// TIA Portal V20 export
// export: Created 2026-10-12T15:48:35.0909134Z, ExportSetting WithDefaults, DisplayName Totally Integrated Automation Portal, DisplayVersion V20, DisplayName TIA Portal Openness, DisplayVersion V20, DisplayName TIA Portal Teamcenter Gateway, DisplayVersion V20, DisplayName TIA Portal Version Control Interface, DisplayVersion V20, DisplayName SINAMICS Startdrive Advanced, DisplayVersion V20 SP1 Update 2, DisplayName SINAMICS Startdrive G110M, G120, G120C, G120D, G120P, G115D, DisplayVersion V20 SP1 Update 2, DisplayName SINAMICS Startdrive G130, G150, S120, S150, SINAMICS MV, G220, S200, S210, DisplayVersion V20 SP1 Update 2, DisplayName STEP 7 Professional, DisplayVersion V20, DisplayName STEP 7 Safety, DisplayVersion V20, DisplayName WinCC Basic/Comfort/Advanced, DisplayVersion V20, DisplayName WinCC Professional, DisplayVersion V20, DisplayName WinCC Unified, DisplayVersion V20
FUNCTION "FRK_Route_DeclarationCell" : Bool   // FC138, SCL
{ S7_Optimized_Access := 'TRUE' }
VERSION : 0.1
// stored: AutoNumber true, IsIECCheckEnabled false, SetENOAutomatically false, UDAEnableTagReadback false
   VAR_INPUT
      Request : "ST_HmiRequest";
   END_VAR
   VAR_IN_OUT
      Module : "FB_DeclarationCell";
      Hal : "ST_DeclarationCellHal";
      Report : "ST_ReleaseReport";
   END_VAR
   VAR_TEMP
      RouteMatched : Bool;
      Index : Int;
   END_VAR
BEGIN

   #FRK_Route_DeclarationCell := FALSE;
   IF NOT "FRK_PathOwned"(OwnerPath := #Module.Status.Name, TargetPath := #Request.TargetPath) THEN
       RETURN;
   END_IF;
   IF #Request.TargetPath = STRING_TO_WSTRING(#Module.Status.Name) THEN
       FOR #Index := 1 TO 16 DO
           #Module.ManConditions[#Index].Used := FALSE;
       END_FOR;
       "FRK_ManualApply"(Core := #Module.Core,
                         Status := #Module.Status,
                         Request := #Request,
                         Commands := #Module.Catalog,
                         Count := #Module.CatalogCount,
                         Conditions := #Module.ManConditions,
                         Report := #Report,
                         Execute := #Module.Execute,
                         Command := #Module.Command,
                         ManualOwned := #Module.ManualOwned);
       #FRK_Route_DeclarationCell := TRUE;
       RETURN;
   END_IF;
   #RouteMatched := "FRK_Route_DeclarationCylinder"(Module := #Module.Clamp, Hal := #Hal.Clamp, Request := #Request, Report := #Report);
   #FRK_Route_DeclarationCell := #FRK_Route_DeclarationCell OR #RouteMatched;
   #RouteMatched := "FRK_Route_DeclarationCylinder"(Module := #Module.Gate, Hal := #Hal.Gate, Request := #Request, Report := #Report);
   #FRK_Route_DeclarationCell := #FRK_Route_DeclarationCell OR #RouteMatched;
END_FUNCTION
